PROGRAM main
  VAR
    S1 AT %IX0.0 : BOOL; (* pulsador NA *)
    H1 AT %QX0.0 : BOOL; (* luz que cambia al apretar *)
    H2 AT %QX0.1 : BOOL; (* luz que cambia al soltar *)
    APRIETA      : R_TRIG;
    SUELTA       : F_TRIG;
    PULSO        : BOOL; (* un ciclo al apretar *)
    PULSO2       : BOOL; (* un ciclo al soltar *)
  END_VAR
  VAR  (* added by the conversion: wires and edge detectors of the diagram *)
    _XOR4_OUT : BOOL;
    _XOR11_OUT : BOOL;
  END_VAR

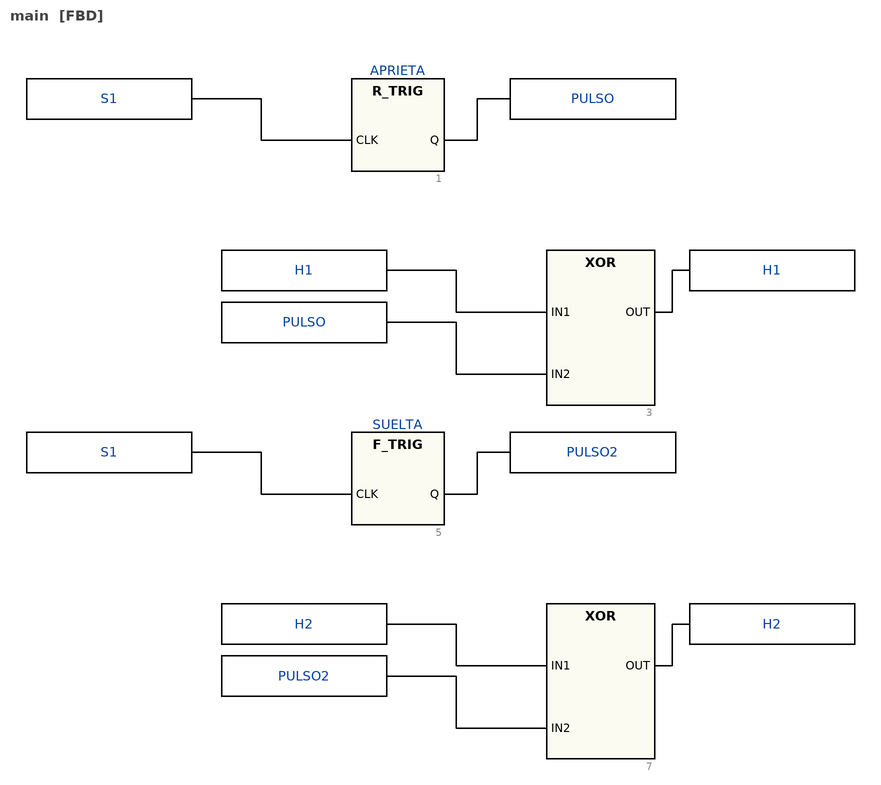
(* FBD diagram, written out as Structured Text *)
APRIETA(CLK := S1);
PULSO := APRIETA.Q;
_XOR4_OUT := H1 XOR PULSO;
H1 := _XOR4_OUT;
SUELTA(CLK := S1);
PULSO2 := SUELTA.Q;
_XOR11_OUT := H2 XOR PULSO2;
H2 := _XOR11_OUT;
END_PROGRAM
